  Folder MAIN
    Script: command_manager(external_control="uGO", cond_suspend=(ITM_Manipulated and AMR_AtTarget and AMR_Charging and AMR_Battery<40), cond_unsuspend=(AMR_Battery≟60))
    Script: log_state(STATE_Info)
    Switch expression=STATE
      Case (caseValue=1)
        Folder Stopping [hidden by the author, left out]
      Case (caseValue=2)
        Folder Stopped [hidden by the author, left out]
      Case (caseValue=3)
        Folder  Resetting [hidden by the author, left out]
      Case (caseValue=4)
        Folder Idle [hidden by the author, left out]
      Case (caseValue=5)
        Folder Starting
          STATE_Info := "Starting"
          'ADD COMMANDS WHAT TO START WITH'
          Call Sub_AMR_MiR_V3
          Folder get ugo data
            Folder Assign Tasks
              Script: TASK.ID = ugo_get_task()
              If TASK.ID≟1
                Task_info := "Charge"
                Folder Parameters [hidden by the author, left out]
              ElseIf TASK.ID≟9
                'Pick Sarstedt Rack from Variable source'
                Task_info := "Navigate to Target"
                Folder Parameters [hidden by the author, left out]
              ElseIf TASK.ID≟13
                Task_info := "Dose Powder"
                Folder Parameters
                  ITM_ID := 1
                  W_now := (UGO.read_input("00","Container_weight"))/1000
                  Pow_name := (UGO.read_input("00","Powder_name"))
                  target_weight := (UGO.read_input("00","Target_weight"))/1000
                  Script: params_init()
                  Script: send_picking_info(Pow_name,target_weight)
                  SuppressedNode
                    w_dosed_total := 0
                  OBJ_Type := 6
                  JIG := 17
                  AMR_PosTarget := 5
              ElseIf TASK.ID≟49
                Task_info := "Pick Containers"
                Folder Parameters
                  ITM_ID := 1
                  OBJ_Type := 6
                  JIG := 15
                  AMR_PosTarget := 3
              ElseIf TASK.ID≟50
                Task_info := "Decap Containers"
                Folder Parameters
                  ITM_ID := 1
                  OBJ_Type := 6
                  JIG := 16
                  AMR_PosTarget := 5
              ElseIf TASK.ID≟51
                Task_info := "Detect Spatula and transfer powder"
                Folder Parameters
                  ITM_ID := 1
                  target_weight := (UGO.read_input("00","Target_weight"))/1000
                  OBJ_Type := 8
                  JIG := 16
                  AMR_PosTarget := 5
              ElseIf TASK.ID≟52
                Task_info := "Pick Powder"
                Folder Parameters
                  ITM_ID := 1
                  SuppressedNode
                    Pow_name := (UGO.read_input("00","Powder_name"))
                  OBJ_Type := 6
                  JIG := 15
                  AMR_PosTarget := 3
              ElseIf TASK.ID≟53
                Task_info := "Decap Powder"
                Folder Parameters
                  ITM_ID := 1
                  OBJ_Type := 6
                  JIG := 1
                  AMR_PosTarget := 5
              ElseIf TASK.ID≟54
                Task_info := "Empty and swap Powder container"
                SuppressedNode
                  Folder Parameters
                    ITM_ID := 1
                    target_weight := (UGO.read_input("00","Target_weight"))/1000
                    W_now := (UGO.read_input("00","Container_weight"))/1000
                    Pow_name := (UGO.read_input("00","Powder_name"))
                    OBJ_Type := 6
                    JIG := 17
                    AMR_PosTarget := 5
                Folder Parameters
                  ITM_ID := 1
                  SuppressedNode
                    target_weight := (UGO.read_input("00","target_weight"))/1000
                  W_now := (UGO.read_input("00","Container_weight"))/1000
                  Pow_name := (UGO.read_input("00","Powder_name"))
                  SuppressedNode
                    Script: scooping_init()
                  SuppressedNode
                    target_weight := W_now-W_EMPTY-(0.002*W_FULL)
                  OBJ_Type := 6
                  JIG := 17
                  AMR_PosTarget := 5
              ElseIf TASK.ID≟55
                Task_info := "Place Powder"
                Folder Parameters
                  ITM_ID := 1
                  OBJ_Type := 6
                  JIG := 21
                  AMR_PosTarget := 5
              ElseIf TASK.ID≟56
                Task_info := "Dose Powder"
                Folder Parameters
                  ITM_ID := 1
                  target_weight := (UGO.read_input("00","Target_weight"))/1000
                  W_now := (UGO.read_input("00","Container_weight"))/1000
                  Pow_name := (UGO.read_input("00","Powder_name"))
                  OBJ_Type := 6
                  JIG := 17
                  AMR_PosTarget := 5
              ElseIf TASK.ID≟57
                Task_info := "Recipe Powder dosing"
                Folder Parameters
                  ITM_ID := 1
                  Pow_A := (UGO.read_input("00","PowderA"))
                  Pow_B := (UGO.read_input("00","PowderB"))
                  Pow_C := (UGO.read_input("00","PowderC"))
                  Total_weight := (UGO.read_input("00","Total_weight"))/1000
                  Pow_A_percent := (UGO.read_input("00","PowderA_percentage"))/100
                  Pow_B_percent := (UGO.read_input("00","PowderB_percentage"))/100
                  Pow_C_percent := (UGO.read_input("00","PowderC_percentage"))/100
                  OBJ_Type := 6
                  JIG := 17
                  AMR_PosTarget := 5
              ElseIf TASK.ID≟58
                Task_info := "Pick Powder containers"
                Folder Parameters [hidden by the author, left out]
              ElseIf TASK.ID≟59
                Task_info := "Empty Powder container"
                Folder Parameters
                  ITM_ID := 1
                  SuppressedNode
                    W_now := (UGO.read_input("00","Container_weight"))/1000
                  Pow_name := (UGO.read_input("00","Powder_name"))
                  SuppressedNode
                    Script: global target_weight = to_str(aa_weight_cont-empty_weight_g)
                  target_weight := (aa_weight_cont-empty_weight_g)*1000
                  W_now := target_weight
                  Script: send_picking_info(Pow_name,target_weight)
                  w_dosed_total := 0
                  OBJ_Type := 6
                  JIG := 17
                  AMR_PosTarget := 5
              ElseIf TASK.ID≟61
                Task_info := "Weigh, Place & Decap"
                Folder Parameters
                  ITM_ID := 1
                  OBJ_Type := 6
                  JIG := 21
                  AMR_PosTarget := 5
              ElseIf TASK.ID≟62
                Task_info := "Dose Powder"
                Folder Parameters
                  ITM_ID := 1
                  SuppressedNode
                    W_now := (UGO.read_input("00","Container_weight"))/1000
                  W_now := aa_weight_cont
                  Pow_name := (UGO.read_input("00","Powder_name"))
                  target_weight := (UGO.read_input("00","Target_weight"))/1000
                  SuppressedNode
                    target_weight := (aa_weight_cont-empty_weight_g)*1000
                  Script: params_init()
                  Script: send_picking_info(Pow_name,target_weight)
                  OBJ_Type := 6
                  JIG := 17
                  AMR_PosTarget := 5
              ElseIf TASK.ID≟63
                Folder Parameters
                  ITM_ID := 1
                  OBJ_Type := 6
                  JIG := 22
                  AMR_PosTarget := 7
              Else 
                Script: set_error(ERROR_WRONG_ORDER)
          Folder test ugo
            Wait Sleep waitTime=0.2
            Script: ugo_update_outputs()
          If starting() and AMR_Done
            Script: log_message(Task_info, "New Task: ")
            Script: log_message(to_str(TASK.ID), "Task_ID: ")
            Script: do_transition(keep_rxry=OBJ_Picked)
            STATE := 6
            Script: ugo_update_outputs()
      Case (caseValue=6)
        Folder Execute
          STATE_Info := "Execute"
          If not CMD_Hold and not CMD_Suspend (checkContinuously=true)
            Switch expression=PROCESS_Step
              Case (caseValue=0)
                PROCESS_Info := "process control"
                Script: log_process(PROCESS_Info)
                Folder process control
                  If not AMR_AtTarget
                    PROCESS_Step := 1
                  ElseIf (( not ITM_Prepared and  not WRK_Done) or (ITM_Prepared and WRK_Done))
                    PROCESS_Step := 2
                  ElseIf not WRK_Done
                    PROCESS_Step := 3
                  Else 
                    Folder task finished
                      PROCESS_Info := ""
                      STATE := 7
                      Script: ugo_update_outputs()
              Case (caseValue=1)
                Folder navigate [hidden by the author, left out]
              Case (caseValue=2)
                Folder prepare
                  'THINGS THAT HAVE TO BE DONE ONCE IN A SEQUENCE,WORKFLOW'
                  PROCESS_Info := "prepare for work"
                  Script: log_process(PROCESS_Info)
                  If TASK.WORK.ITM_ID_Src>1
                    ITM_ID := TASK.WORK.ITM_ID_Src
                  ElseIf TASK.WORK.ITM_ID_Tgt>1
                    ITM_ID := TASK.WORK.ITM_ID_Tgt
                  If not ARM_Referenced and (ITM_ID≠0)
                    STP := 1
                  ElseIf ARM_Referenced or (ITM_ID≟0)
                    STP := 2
                  Switch expression=STP
                    Case (caseValue=1)
                      Folder reference [hidden by the author, left out]
                    Case (caseValue=2)
                      Folder manipulate [hidden by the author, left out]
                  ITM_Prepared := (ITM_Manipulated or  not found_in_list(ITM_ID, ITM_ID_List)) and (ARM_Referenced or ITM_ID≟0) and  not WRK_Done
                  STP := 0
                  STP_Info := ""
                  PROCESS_Step := 0
              Case (caseValue=3)
                Folder work
                  'ADD EVERY MACHINE, OBJECT, STATION TO WORK ON'
                  Switch expression=ITM_ID
                    Case (caseValue=1)
                      Folder uLM
                        If TASK.ID≟12
                          Folder fill racks [hidden by the author, left out]
                        ElseIf TASK.ID≟13
                          Folder Dose Powder
                            Action := 131
                            Call Sub_Vision_V18
                            Action := 34
                            Call Sub_Action_V4
                            PROCESS_Step := 0
                            WRK_Done := True
                        ElseIf TASK.ID≟49
                          Folder Pick Powder container [hidden by the author, left out]
                        ElseIf TASK.ID≟50
                          Folder Decap containers [hidden by the author, left out]
                        ElseIf TASK.ID≟51
                          Folder Detect Spatula and transfer powder [hidden by the author, left out]
                        ElseIf TASK.ID≟52
                          Folder Pick Powder container
                            Action := 131
                            Call Sub_Vision_V18
                            Action := 39
                            Call Sub_Action_V4
                            PROCESS_Step := 0
                            WRK_Done := True
                        ElseIf TASK.ID≟53
                          Folder Decap containerA
                            Action := 40
                            Call Sub_Action_V4
                            PROCESS_Step := 0
                            WRK_Done := True
                        ElseIf TASK.ID≟55
                          Folder Place Powder
                            Action := 131
                            Call Sub_Vision_V18
                            Action := 41
                            Call Sub_Action_V4
                            PROCESS_Step := 0
                            WRK_Done := True
                        ElseIf TASK.ID≟54
                          Folder Empty and swap container
                            Action := 131
                            Call Sub_Vision_V18
                            Action := 42
                            Call Sub_Action_V4
                            PROCESS_Step := 0
                            WRK_Done := True
                        ElseIf TASK.ID≟56
                          Folder Dispense Powder [hidden by the author, left out]
                        ElseIf TASK.ID≟57
                          Folder Recipe Dosing
                            Action := 48
                            Call Sub_Action_V4
                            SuppressedNode
                              Script: recipe_init(Pow_A, Pow_B, Pow_C, Total_weight, Pow_A_percent, Pow_B_percent, Pow_C_percent)
                            SuppressedNode
                              Loop While (checkContinuously=false) expression=recipe_next()≟ True
                                Action := 44
                                Call Sub_Action_V4
                                JIG := 21
                                Action := 131
                                Call Sub_Vision_V18
                                Action := 45
                                Call Sub_Action_V4
                                Script: dosing_start()
                                JIG := 17
                                Action := 131
                                Call Sub_Vision_V18
                                Action := 46
                                Call Sub_Action_V4
                                Script: dosing_end()
                            PROCESS_Step := 0
                            WRK_Done := True
                        ElseIf TASK.ID≟58
                          Folder Pick Powder containers
                            Num_cont_picked := 0
                            powder_position := "Position1"
                            Loop While (checkContinuously=false) expression=Num_cont_picked<3
                              Action := 131
                              Call Sub_Vision_V18
                              Action := 47
                              Call Sub_Action_V4
                            PROCESS_Step := 0
                            WRK_Done := True
                        ElseIf TASK.ID≟59
                          Folder Empty powder container
                            Action := 131
                            Call Sub_Vision_V18
                            Action := 50
                            Call Sub_Action_V4
                            PROCESS_Step := 0
                            WRK_Done := True
                        ElseIf TASK.ID≟61
                          Folder Place Powder
                            Action := 131
                            Call Sub_Vision_V18
                            Action := 51
                            Call Sub_Action_V4
                            PROCESS_Step := 0
                            WRK_Done := True
                        ElseIf TASK.ID≟62
                          Folder Dose Powder [hidden by the author, left out]
                        ElseIf TASK.ID≟63
                          Folder Swabbing
                            Action := 131
                            Call Sub_Vision_V18
                            Action := 53
                            Call Sub_Action_V4
                            SuppressedNode
                              Action := 55
                            SuppressedNode
                              Call Sub_Action_V4
                            PROCESS_Step := 0
                            WRK_Done := True
                    Case (caseValue=2)
                      SuppressedNode
                        Folder Centrfiuge
                          SuppressedNode
                            Script: cent_error_check()
                          OBJ_Type := 1
                          If not ERROR.FLAG
                            'load racks'
                            If TASK.ID≟14
                              Loop While (checkContinuously=false) expression=(PRC_RackCounter<4) and  not CMD_Stop and  not ERROR.FLAG
                                ITM_ID := TASK.WORK.ITM_ID_Src
                                JIG := 4
                                JIG_Slot := PRC_RackCounter+1
                                Action := 1
                                CallSubProgram
                                If OBJ_Picked and  not ERROR.FLAG
                                  ITM_ID := TASK.WORK.ITM_ID_Tgt
                                  Script: execute_cent_action(ACTION_ROTATE, JIG_Slot)
                                  Action := 7
                                  CallSubProgram
                                  PRC_RackCounter := PRC_RackCounter + 1
                              If not ERROR.FLAG
                                WRK_Done := True
                                PROCESS_Step := 0
                            'unload racks'
                            If TASK.ID≟15
                              If CNT_State_Actual≟2 or CNT_State_Actual≟3
                                Loop While (checkContinuously=false) expression=(PRC_RackCounter<4) and  not CMD_Stop and  not ERROR.FLAG
                                  ITM_ID := TASK.WORK.ITM_ID_Src
                                  JIG_Slot := PRC_RackCounter + 1
                                  Script: execute_cent_action(ACTION_ROTATE, JIG_Slot)
                                  Script: execute_cent_action(ACTION_INSPECT, JIG_Slot)
                                  Action := 8
                                  CallSubProgram
                                  If OBJ_Picked and  not ERROR.FLAG
                                    ITM_ID := TASK.WORK.ITM_ID_Tgt
                                    JIG := 4
                                    JIG_Slot := PRC_RackCounter + 1
                                    Action := 2
                                    CallSubProgram
                                    PRC_RackCounter := PRC_RackCounter+1
                                If not ERROR.FLAG
                                  WRK_Done := True
                                  PROCESS_Step := 0
                    Case (caseValue=5)
                      SuppressedNode
                        Folder SarstedtTable
                          Action := 131
                          CallSubProgram
                          Action := 1
                          CallSubProgram
                          PROCESS_Step := 0
                          WRK_Done := True
                    Case (caseValue=20)
                      SuppressedNode
                        Folder Biorad rack
                          'load racks'
                          If Task_ID≟16
                            SuppressedNode
                              PRC_RackCounter := 0
                            Loop While (checkContinuously=false) expression=(PRC_RackCounter<PRC_RackNumber) and  not CMD_Stop
                              JIG_Slot := PRC_RackCounter
                              Action := 1
                              PRC_Target := 0
                              CallSubProgram
                              If OBJ_Picked
                                Action := 2
                                PRC_Target := 1
                                CallSubProgram
                                Action := 7
                                PRC_Target := 1
                                CallSubProgram
                                PRC_RackCounter := PRC_RackCounter+1
                            WRK_Done := True
                            PROCESS_Step := 0
                          'unload racks'
                          SuppressedNode
                            If Task_ID≟17
                              SuppressedNode
                                PRC_RackCounter := 0
                              Loop While (checkContinuously=false) expression=(PRC_RackCounter<PRC_RackNumber) and  not CMD_Stop
                                JIG_Slot := PRC_RackCounter
                                Action := 8
                                PRC_Target := 1
                                Script: textmsg("Callactionunload=",Action)
                                CallSubProgram
                                Action := 1
                                PRC_Target := 1
                                Script: textmsg("Callactionpick=",Action)
                                CallSubProgram
                                If OBJ_Picked
                                  Action := 2
                                  PRC_Target := 0
                                  Script: textmsg("Callactionplace=",Action)
                                  CallSubProgram
                                  PRC_RackCounter := PRC_RackCounter+1
                              WRK_Done := True
                              PROCESS_Step := 0
                          If Task_ID≟17
                            PRC_RackCounter := 0
                            Loop While (checkContinuously=false) expression=(PRC_RackCounter<PRC_RackNumber) and  not CMD_Stop
                              Wait Condition expression=SensorData[PRC_RackCounter]≟1
                              JIG_Slot := PRC_RackCounter
                              Action := 8
                              PRC_Target := 1
                              Script: textmsg("Callactionunload=",Action)
                              CallSubProgram
                              Action := 1
                              PRC_Target := 1
                              Script: textmsg("Callactionpick=",Action)
                              CallSubProgram
                              If OBJ_Picked
                                Action := 2
                                PRC_Target := 0
                                Script: textmsg("Callactionplace=",Action)
                                CallSubProgram
                                PRC_RackCounter := PRC_RackCounter+1
                            WRK_Done := True
                            PROCESS_Step := 0
                    Case (caseValue=43)
                      SuppressedNode
                        Folder Pick the rack
                          Action := 131
                          CallSubProgram
                          Action := 1
                          CallSubProgram
                          PROCESS_Step := 0
                          WRK_Done := True
                    Case (caseValue=2147483647)
                      WRK_Done := True
                      PROCESS_Step := 0
          If CMD_Hold
            STATE := 9
            Script: ugo_update_outputs()
          ElseIf CMD_Suspend
            STATE := 12
            Script: ugo_update_outputs()
      Case (caseValue=7)
        Folder Completing [hidden by the author, left out]
      Case (caseValue=8)
        Folder Complete [hidden by the author, left out]
      Case (caseValue=9)
        Folder Holding [hidden by the author, left out]
      Case (caseValue=10)
        Folder Held [hidden by the author, left out]
      Case (caseValue=11)
        Folder Unholding [hidden by the author, left out]
      Case (caseValue=12)
        Folder Suspending [hidden by the author, left out]
      Case (caseValue=13)
        Folder Suspended [hidden by the author, left out]
      Case (caseValue=14)
        Folder Unsuspending [hidden by the author, left out]
      Case (caseValue=15)
        Folder Aborting [hidden by the author, left out]
      Case (caseValue=16)
        Folder Aborted [hidden by the author, left out]
      Case (caseValue=17)
        Folder Clearing [hidden by the author, left out]
    Script: log_state(STATE_Info)
    Script: log_warning(WARNING.MSG)
    Script: log_error(ERROR.MSG)
    Folder Times [hidden by the author, left out]
    SuppressedNode
      Script: sync()
    Wait Sleep waitTime=0.1
Thread Thread_1 (runOnlyOnce=false)
  Folder Dosing Weight [hidden by the author, left out]
  Script: sync()
Thread Thread_2 (runOnlyOnce=false)
  Folder Vibration motor [hidden by the author, left out]
  Script: sync()
Thread Thread_3 (runOnlyOnce=false)
  Folder Container weight [hidden by the author, left out]
  Script: sync()
SubProgram -> Sub_Vision_V18
SubProgram  [hidden by the author, left out]
SubProgram -> Sub_Action_V4
